// TIA Portal V20 export
// export: Created 2026-10-12T04:58:24.2013317Z, ExportSetting WithDefaults, DisplayName Totally Integrated Automation Portal, DisplayVersion V20, DisplayName TIA Portal Openness, DisplayVersion V20, DisplayName TIA Portal Teamcenter Gateway, DisplayVersion V20, DisplayName TIA Portal Version Control Interface, DisplayVersion V20, DisplayName SINAMICS Startdrive Advanced, DisplayVersion V20 SP1 Update 2, DisplayName SINAMICS Startdrive G110M, G120, G120C, G120D, G120P, G115D, DisplayVersion V20 SP1 Update 2, DisplayName SINAMICS Startdrive G130, G150, S120, S150, SINAMICS MV, G220, S200, S210, DisplayVersion V20 SP1 Update 2, DisplayName STEP 7 Professional, DisplayVersion V20, DisplayName STEP 7 Safety, DisplayVersion V20, DisplayName WinCC Basic/Comfort/Advanced, DisplayVersion V20, DisplayName WinCC Professional, DisplayVersion V20, DisplayName WinCC Unified, DisplayVersion V20
FUNCTION "FRK_CfgWrite_SatelliteUnit" : Bool   // FC151, SCL
{ S7_Optimized_Access := 'TRUE' }
VERSION : 0.1
// stored: AutoNumber true, IsIECCheckEnabled false, SetENOAutomatically false, UDAEnableTagReadback false
   VAR_INPUT
      Request : "ST_HmiRequest";
      Access : "FRK_Access";
      RootIndex : Int;
      RootReady : Bool;
   END_VAR
   VAR_IN_OUT
      Module : "FB_SatelliteUnit";
      Matched : Bool;
   END_VAR
   VAR_TEMP
      Ok : Bool;
      Level : DInt;
      Code : String[64];
      Inactive : Bool;
   END_VAR
BEGIN

   #FRK_CfgWrite_SatelliteUnit := FALSE;
   IF #Request.TargetPath = STRING_TO_WSTRING(#Module.Status.Name) OR (#Request.TargetPath = WSTRING#'' AND #Module.Core.ParentIndex = 0) THEN
       "FRK_CfgDef_SatelliteUnit"(FieldIndex := 1);
       IF #Request.NameValue = "FRK_ConfigScratch".Entry.WriteKey THEN
           #Matched := TRUE;
           IF DINT_TO_UDINT(#Request.IntValue) <> "FRK_ConfigScratch".Entry.WriteRevision THEN
               RETURN;
           END_IF;
           #Level := MAX(IN1 := #Access.Policy.Required[1], IN2 := "FRK_ConfigScratch".MinWrite);
           IF #Access.CurrentLevel < #Level THEN
               RETURN;
           END_IF;
           IF #Request.DurationMs <> 0 THEN
               RETURN;
           END_IF;
           #Code := "FRK_ConfigModelCode"(RootIndex := #RootIndex, ModelIndex := #Request.DurationMs);
           #Inactive := #Code <> "FRK_ConfigStore".ActiveModels[#RootIndex];
           IF "FRK_ConfigScratch".Entry.RequiresReady AND NOT #Inactive AND NOT #RootReady THEN
               RETURN;
           END_IF;
           #Ok := "FRK_ConfigDecode"(Text := #Request.TextValue, Storage := "FRK_ConfigScratch".Storage, Minimum := "FRK_ConfigScratch".Minimum, Maximum := "FRK_ConfigScratch".Maximum, MaxLength := "FRK_ConfigScratch".MaxLength, Value := "FRK_ConfigScratch".Value);
           IF NOT #Ok THEN
               RETURN;
           END_IF;
           #Ok := "FRK_ConfigPut"(Scope := #Module.Status.Name, ModelCode := #Code, Text := #Request.TextValue, RootIndex := #RootIndex);
           IF NOT #Ok THEN
               RETURN;
           END_IF;
           IF NOT #Inactive THEN
               #Module.ParCfg.Timeout := DINT_TO_TIME(LINT_TO_DINT("FRK_ConfigScratch".Value.Number));
           END_IF;
           #FRK_CfgWrite_SatelliteUnit := TRUE;
           RETURN;
       END_IF;
       "FRK_CfgDef_SatelliteUnit"(FieldIndex := 2);
       IF #Request.NameValue = "FRK_ConfigScratch".Entry.WriteKey THEN
           #Matched := TRUE;
           IF DINT_TO_UDINT(#Request.IntValue) <> "FRK_ConfigScratch".Entry.WriteRevision THEN
               RETURN;
           END_IF;
           #Level := MAX(IN1 := #Access.Policy.Required[1], IN2 := "FRK_ConfigScratch".MinWrite);
           IF #Access.CurrentLevel < #Level THEN
               RETURN;
           END_IF;
           IF #Request.DurationMs <> 0 THEN
               RETURN;
           END_IF;
           #Code := "FRK_ConfigModelCode"(RootIndex := #RootIndex, ModelIndex := #Request.DurationMs);
           #Inactive := #Code <> "FRK_ConfigStore".ActiveModels[#RootIndex];
           IF "FRK_ConfigScratch".Entry.RequiresReady AND NOT #Inactive AND NOT #RootReady THEN
               RETURN;
           END_IF;
           #Ok := "FRK_ConfigDecode"(Text := #Request.TextValue, Storage := "FRK_ConfigScratch".Storage, Minimum := "FRK_ConfigScratch".Minimum, Maximum := "FRK_ConfigScratch".Maximum, MaxLength := "FRK_ConfigScratch".MaxLength, Value := "FRK_ConfigScratch".Value);
           IF NOT #Ok THEN
               RETURN;
           END_IF;
           #Ok := "FRK_ConfigPut"(Scope := #Module.Status.Name, ModelCode := #Code, Text := #Request.TextValue, RootIndex := #RootIndex);
           IF NOT #Ok THEN
               RETURN;
           END_IF;
           IF NOT #Inactive THEN
               #Module.ParCfg.Preset := LINT_TO_DINT("FRK_ConfigScratch".Value.Number);
           END_IF;
           #FRK_CfgWrite_SatelliteUnit := TRUE;
           RETURN;
       END_IF;
       "FRK_CfgDef_SatelliteUnit"(FieldIndex := 3);
       IF #Request.NameValue = "FRK_ConfigScratch".Entry.WriteKey THEN
           #Matched := TRUE;
           IF DINT_TO_UDINT(#Request.IntValue) <> "FRK_ConfigScratch".Entry.WriteRevision THEN
               RETURN;
           END_IF;
           #Level := MAX(IN1 := #Access.Policy.Required[1], IN2 := "FRK_ConfigScratch".MinWrite);
           IF #Access.CurrentLevel < #Level THEN
               RETURN;
           END_IF;
           IF #Request.DurationMs <> 0 THEN
               RETURN;
           END_IF;
           #Code := '';
           #Inactive := FALSE;
           IF "FRK_ConfigScratch".Entry.RequiresReady AND NOT #Inactive AND NOT #RootReady THEN
               RETURN;
           END_IF;
           #Ok := "FRK_ConfigDecode"(Text := #Request.TextValue, Storage := "FRK_ConfigScratch".Storage, Minimum := "FRK_ConfigScratch".Minimum, Maximum := "FRK_ConfigScratch".Maximum, MaxLength := "FRK_ConfigScratch".MaxLength, Value := "FRK_ConfigScratch".Value);
           IF NOT #Ok THEN
               RETURN;
           END_IF;
           #Ok := "FRK_ConfigPut"(Scope := #Module.Status.Name, ModelCode := #Code, Text := #Request.TextValue, RootIndex := #RootIndex);
           IF NOT #Ok THEN
               RETURN;
           END_IF;
           IF NOT #Inactive THEN
               #Module.StationCfg.SiteLabel := "FRK_ConfigScratch".Value.Text;
           END_IF;
           #FRK_CfgWrite_SatelliteUnit := TRUE;
           RETURN;
       END_IF;
       "FRK_CfgDef_SatelliteUnit"(FieldIndex := 4);
       IF #Request.NameValue = "FRK_ConfigScratch".Entry.WriteKey THEN
           #Matched := TRUE;
           IF DINT_TO_UDINT(#Request.IntValue) <> "FRK_ConfigScratch".Entry.WriteRevision THEN
               RETURN;
           END_IF;
           #Level := MAX(IN1 := #Access.Policy.Required[1], IN2 := "FRK_ConfigScratch".MinWrite);
           IF #Access.CurrentLevel < #Level THEN
               RETURN;
           END_IF;
           IF #Request.DurationMs <> 0 THEN
               RETURN;
           END_IF;
           #Code := '';
           #Inactive := FALSE;
           IF "FRK_ConfigScratch".Entry.RequiresReady AND NOT #Inactive AND NOT #RootReady THEN
               RETURN;
           END_IF;
           #Ok := "FRK_ConfigDecode"(Text := #Request.TextValue, Storage := "FRK_ConfigScratch".Storage, Minimum := "FRK_ConfigScratch".Minimum, Maximum := "FRK_ConfigScratch".Maximum, MaxLength := "FRK_ConfigScratch".MaxLength, Value := "FRK_ConfigScratch".Value);
           IF NOT #Ok THEN
               RETURN;
           END_IF;
           #Ok := "FRK_ConfigPut"(Scope := #Module.Status.Name, ModelCode := #Code, Text := #Request.TextValue, RootIndex := #RootIndex);
           IF NOT #Ok THEN
               RETURN;
           END_IF;
           IF NOT #Inactive THEN
               #Module.StationCfg.LongText := "FRK_ConfigScratch".Value.Text;
           END_IF;
           #FRK_CfgWrite_SatelliteUnit := TRUE;
           RETURN;
       END_IF;
       "FRK_CfgDef_SatelliteUnit"(FieldIndex := 5);
       IF #Request.NameValue = "FRK_ConfigScratch".Entry.WriteKey THEN
           #Matched := TRUE;
           IF DINT_TO_UDINT(#Request.IntValue) <> "FRK_ConfigScratch".Entry.WriteRevision THEN
               RETURN;
           END_IF;
           #Level := MAX(IN1 := #Access.Policy.Required[1], IN2 := "FRK_ConfigScratch".MinWrite);
           IF #Access.CurrentLevel < #Level THEN
               RETURN;
           END_IF;
           IF #Request.DurationMs <> 0 THEN
               RETURN;
           END_IF;
           #Code := '';
           #Inactive := FALSE;
           IF "FRK_ConfigScratch".Entry.RequiresReady AND NOT #Inactive AND NOT #RootReady THEN
               RETURN;
           END_IF;
           #Ok := "FRK_ConfigDecode"(Text := #Request.TextValue, Storage := "FRK_ConfigScratch".Storage, Minimum := "FRK_ConfigScratch".Minimum, Maximum := "FRK_ConfigScratch".Maximum, MaxLength := "FRK_ConfigScratch".MaxLength, Value := "FRK_ConfigScratch".Value);
           IF NOT #Ok THEN
               RETURN;
           END_IF;
           #Ok := "FRK_ConfigPut"(Scope := #Module.Status.Name, ModelCode := #Code, Text := #Request.TextValue, RootIndex := #RootIndex);
           IF NOT #Ok THEN
               RETURN;
           END_IF;
           IF NOT #Inactive THEN
               #Module.StationCfg.Enabled := "FRK_ConfigScratch".Value.Flag;
           END_IF;
           #FRK_CfgWrite_SatelliteUnit := TRUE;
           RETURN;
       END_IF;
   END_IF;
   #Ok := "FRK_CfgWrite_DeclarationCell"(Module := #Module.Cell, Access := #Access, Request := #Request, RootIndex := #RootIndex, RootReady := #RootReady, Matched := #Matched);
   IF #Matched THEN
       #FRK_CfgWrite_SatelliteUnit := #Ok;
       RETURN;
   END_IF;
   #Ok := "FRK_CfgWrite_InnerUnit"(Module := #Module.Inner, Access := #Access, Request := #Request, RootIndex := #RootIndex, RootReady := #RootReady, Matched := #Matched);
   IF #Matched THEN
       #FRK_CfgWrite_SatelliteUnit := #Ok;
       RETURN;
   END_IF;
END_FUNCTION
